// TIA Portal V20 export
// export: Created 2026-10-11T05:28:40.709762Z, ExportSetting WithDefaults, DisplayName Totally Integrated Automation Portal, DisplayVersion V20, DisplayName TIA Portal Openness, DisplayVersion V20, DisplayName TIA Portal Teamcenter Gateway, DisplayVersion V20, DisplayName TIA Portal Version Control Interface, DisplayVersion V20, DisplayName SINAMICS Startdrive Advanced, DisplayVersion V20 SP1 Update 2, DisplayName SINAMICS Startdrive G110M, G120, G120C, G120D, G120P, G115D, DisplayVersion V20 SP1 Update 2, DisplayName SINAMICS Startdrive G130, G150, S120, S150, SINAMICS MV, G220, S200, S210, DisplayVersion V20 SP1 Update 2, DisplayName STEP 7 Professional, DisplayVersion V20, DisplayName STEP 7 Safety, DisplayVersion V20, DisplayName WinCC Basic/Comfort/Advanced, DisplayVersion V20, DisplayName WinCC Professional, DisplayVersion V20, DisplayName WinCC Unified, DisplayVersion V20
FUNCTION "FRK_UnitRunStart" : Void   // FC48, SCL
{ S7_Optimized_Access := 'TRUE' }
VERSION : 0.1
// stored: AutoNumber true, IsIECCheckEnabled false, SetENOAutomatically false, UDAEnableTagReadback false
   VAR_INPUT
      Timeout : Time;
      Label : String;
   END_VAR
   VAR_IN_OUT
      Core : "FRK_Core";
      Status : "ST_ModuleStatus";
   END_VAR
BEGIN

   "FRK_Start"(Core := #Core,
               Status := #Status,
               Supported := TRUE,
               Timeout := #Timeout,
               Label := #Label);
   // A continuous run ends at Stop. Bounded commands/steps own progress timeouts.
   #Core.TimeoutMs := 0;
END_FUNCTION
